DATA_BLOCK "DI_SYSTEM_STRING_NAMES_ENG"
{ S7_Optimized_Access := 'FALSE' }
VERSION : 0.1
NON_RETAIN
"DT_DI_STRING_SYSTEM_NAMES"

BEGIN
   NUM[0] := 'Unit control and prot. +1CJA01';
   NUM[1] := 'Unit control and prot. +1CJA01';
   NUM[2] := 'Unit control and prot. +1CJA01';
   NUM[3] := 'Unit control and prot. +1CJA01';
   NUM[4] := 'Unit control and prot. +1CJA01';
   NUM[5] := 'Unit control and prot. +1CJA01';
   NUM[6] := 'Unit control and prot. +1CJA01';
   NUM[7] := 'Power house pushbutton ';
   NUM[8] := 'Unit control and prot. +1CJA01';
   NUM[9] := '';
   NUM[10] := 'Unit control and prot. +1CJA01';
   NUM[11] := 'Unit control and prot. +1CJA01';
   NUM[12] := 'Unit control and prot. +1CJA01';
   NUM[13] := 'Unit control and prot. +1CJA01';
   NUM[14] := 'Unit control and prot. +1CJA01';
   NUM[15] := '';
   NUM[16] := '';
   NUM[17] := 'Unit GCB cubicle +BAC01';
   NUM[18] := 'Unit GCB cubicle +BAC01';
   NUM[19] := 'Unit GCB cubicle +BAC01';
   NUM[20] := 'Unit GCB cubicle +BAC01';
   NUM[21] := '';
   NUM[22] := '';
   NUM[23] := 'Unit GCB cubicle +BAC01';
   NUM[24] := 'Unit GCB cubicle +BAC01';
   NUM[25] := 'Unit control and prot. +1CJA01';
   NUM[26] := '';
   NUM[27] := '';
   NUM[28] := 'Unit control and prot. +1CJA01';
   NUM[29] := '';
   NUM[30] := 'Unit GCB cubicle +BAC01';
   NUM[31] := 'Common control and prot. +0CJA01';
   NUM[32] := '';
   NUM[33] := '';
   NUM[34] := 'Auxiliary supply cubicle +0BFA01';
   NUM[35] := '';
   NUM[36] := 'Unit Aux. Power Supply +BFA01';
   NUM[37] := '';
   NUM[38] := '';
   NUM[39] := '';
   NUM[40] := '';
   NUM[41] := '';
   NUM[42] := '';
   NUM[43] := '';
   NUM[44] := '';
   NUM[45] := '';
   NUM[46] := '';
   NUM[47] := 'Unit Aux. Power Supply +BFA01';
   NUM[48] := '';
   NUM[49] := 'Unit Aux. Power Supply +BFA01';
   NUM[50] := 'Unit Aux. Power Supply +BFA01';
   NUM[51] := 'Unit Aux. Power Supply +BFA01';
   NUM[52] := '';
   NUM[53] := 'Unit Aux. Power Supply +BFA01';
   NUM[54] := '';
   NUM[55] := '';
   NUM[56] := 'Unit Aux. Power Supply +BFA01';
   NUM[57] := '';
   NUM[58] := 'Unit Aux. Power Supply +BFA01';
   NUM[59] := 'Unit Aux. Power Supply +BFA01';
   NUM[60] := 'Unit Aux. Power Supply +BFA01';
   NUM[61] := 'Unit Aux. Power Supply +BFA01';
   NUM[62] := 'Unit Aux. Power Supply +BFA01';
   NUM[63] := '';
   NUM[64] := '';
   NUM[65] := '';
   NUM[66] := '';
   NUM[67] := '';
   NUM[68] := 'Unit GCB cubicle +BAC01';
   NUM[69] := 'Unit GCB cubicle +BAC01';
   NUM[70] := '';
   NUM[71] := '';
   NUM[72] := '';
   NUM[73] := '';
   NUM[74] := 'Unit GCB cubicle +BAC01';
   NUM[75] := '';
   NUM[76] := '';
   NUM[77] := '';
   NUM[78] := '';
   NUM[79] := '';
   NUM[80] := '';
   NUM[81] := '';
   NUM[82] := '';
   NUM[83] := 'Unit GCB cubicle +BAC01';
   NUM[84] := '';
   NUM[85] := '';
   NUM[86] := 'Unit GCB cubicle +BAC01';
   NUM[87] := '';
   NUM[88] := '';
   NUM[89] := '';
   NUM[90] := '';
   NUM[91] := '';
   NUM[92] := '';
   NUM[93] := '';
   NUM[94] := '';
   NUM[95] := '';
   NUM[96] := '';
   NUM[97] := '';
   NUM[98] := '';
   NUM[99] := 'Unit control and prot. +1CJA01';
   NUM[100] := 'Unit control and prot. +1CJA01';
   NUM[101] := '';
   NUM[102] := '';
   NUM[103] := '';
   NUM[104] := '';
   NUM[105] := '';
   NUM[106] := '';
   NUM[107] := '';
   NUM[108] := '';
   NUM[109] := '';
   NUM[110] := '';
   NUM[111] := '';
   NUM[112] := '';
   NUM[113] := 'Unit Generator - 1MKA10';
   NUM[114] := 'Unit Generator - 1MKA10';
   NUM[115] := '';
   NUM[116] := '';
   NUM[117] := '';
   NUM[118] := '';
   NUM[119] := '';
   NUM[120] := '';
   NUM[121] := '';
   NUM[122] := '';
   NUM[123] := '';
   NUM[124] := '';
   NUM[125] := '';
   NUM[126] := '';
   NUM[127] := '';
   NUM[128] := 'Unit GCB cubicle +BAC01';
   NUM[129] := '';
   NUM[130] := 'Unit GCB cubicle +BAC01';
   NUM[131] := 'Unit GCB cubicle +BAC01';
   NUM[132] := '';
   NUM[133] := '';
   NUM[134] := '';
   NUM[135] := '';
   NUM[136] := '';
   NUM[137] := '';
   NUM[138] := '';
   NUM[139] := '';
   NUM[140] := 'AJA03 - Transformator fedder';
   NUM[141] := '';
   NUM[142] := '';
   NUM[143] := '';
   NUM[144] := '';
   NUM[145] := '';
   NUM[146] := '';
   NUM[147] := '';
   NUM[148] := '';
   NUM[149] := '';
   NUM[150] := '';
   NUM[151] := '';
   NUM[152] := '';
   NUM[153] := '';
   NUM[154] := '';
   NUM[155] := '';
   NUM[156] := '';
   NUM[157] := '';
   NUM[158] := '';
   NUM[159] := '';
   NUM[160] := '';
   NUM[161] := '';
   NUM[162] := '';
   NUM[163] := '';
   NUM[164] := '';
   NUM[165] := '';
   NUM[166] := '';
   NUM[167] := '';
   NUM[168] := '';
   NUM[169] := '';
   NUM[170] := '';
   NUM[171] := '';
   NUM[172] := '';
   NUM[173] := '';
   NUM[174] := '';
   NUM[175] := '';
   NUM[176] := '';
   NUM[177] := '';
   NUM[178] := '';
   NUM[179] := '';
   NUM[180] := '';
   NUM[181] := '';
   NUM[182] := '';
   NUM[183] := '';
   NUM[184] := '';
   NUM[185] := '';
   NUM[186] := '';
   NUM[187] := '';
   NUM[188] := '';
   NUM[189] := '';
   NUM[190] := '';
   NUM[191] := '';
   NUM[192] := 'Unit MIV +1MEA10';
   NUM[193] := '';
   NUM[194] := 'Unit MIV +1MEA10';
   NUM[195] := '';
   NUM[196] := '';
   NUM[197] := '';
   NUM[198] := '';
   NUM[199] := '';
   NUM[200] := '';
   NUM[201] := 'Unit Turbine +1MEA10';
   NUM[202] := 'Unit Turbine +1MEA10';
   NUM[203] := 'Unit control and prot. +1CJA01';
   NUM[204] := '';
   NUM[205] := '';
   NUM[206] := 'Unit control and prot. +1CJA01';
   NUM[207] := 'Unit control and prot. +1CJA01';
   NUM[208] := 'Unit control and prot. +1CJA01';
   NUM[209] := '';
   NUM[210] := '';
   NUM[211] := '';
   NUM[212] := '';
   NUM[213] := '';
   NUM[214] := '';
   NUM[215] := '';
   NUM[216] := '';
   NUM[217] := '';
   NUM[218] := '';
   NUM[219] := '';
   NUM[220] := '';
   NUM[221] := '';
   NUM[222] := '';
   NUM[223] := '';
   NUM[224] := '';
   NUM[225] := 'Unit HPU +1MEX10';
   NUM[226] := '';
   NUM[227] := '';
   NUM[228] := 'Unit HPU +1MEX10';
   NUM[229] := '';
   NUM[230] := '';
   NUM[231] := '';
   NUM[232] := '';
   NUM[233] := 'Unit HPU +1MEX10';
   NUM[234] := 'Unit HPU +1MEX10';
   NUM[235] := '';
   NUM[236] := '';
   NUM[237] := 'Unit HPU +1MEX10';
   NUM[238] := 'Unit HPU +1MEX10';
   NUM[239] := '';
   NUM[240] := '';
   NUM[241] := '';
   NUM[242] := 'Unit control and prot. +1CJA01';
   NUM[243] := 'Unit control and prot. +1CJA01';
   NUM[244] := '';
   NUM[245] := 'HPU +1MEX10';
   NUM[246] := '';
   NUM[247] := '';
   NUM[248] := '';
   NUM[249] := '';
   NUM[250] := '';
   NUM[251] := '';
   NUM[252] := '';
   NUM[253] := '';
   NUM[254] := '';
   NUM[255] := '';
   NUM[256] := '';
   NUM[257] := '';
   NUM[258] := '';
   NUM[259] := 'Unit control and prot. +1CJA01';
   NUM[260] := 'Unit control and prot. +1CJA01';
   NUM[261] := '';
   NUM[262] := '';
   NUM[263] := '';
   NUM[264] := 'Unit control and prot. +1CJA01';
   NUM[265] := 'Unit control and prot. +1CJA01';
   NUM[266] := '';
   NUM[267] := '';
   NUM[268] := '';
   NUM[269] := '';
   NUM[270] := '';
   NUM[271] := '';
   NUM[272] := '';
   NUM[273] := '';
   NUM[274] := '';
   NUM[275] := '';
   NUM[276] := '';
   NUM[277] := '';
   NUM[278] := '';
   NUM[279] := '';
   NUM[280] := '';
   NUM[281] := '';
   NUM[282] := '';
   NUM[283] := '';
   NUM[284] := '';
   NUM[285] := '';
   NUM[286] := '';
   NUM[287] := '';
   NUM[288] := '';
   NUM[289] := '';
   NUM[290] := '';
   NUM[291] := '';
   NUM[292] := '';
   NUM[293] := '';
   NUM[294] := '';
   NUM[295] := '';
   NUM[296] := '';
   NUM[297] := '';
   NUM[298] := '';
   NUM[299] := '';
   NUM[300] := '';
   NUM[301] := '';
   NUM[302] := '';
   NUM[303] := '';
   NUM[304] := '';
   NUM[305] := '';
   NUM[306] := '';
   NUM[307] := '';
   NUM[308] := '';
   NUM[309] := '';
   NUM[310] := '';
   NUM[311] := '';
   NUM[312] := '';
   NUM[313] := '';
   NUM[314] := '';
   NUM[315] := '';
   NUM[316] := '';
   NUM[317] := '';
   NUM[318] := '';
   NUM[319] := '';
   NUM[320] := '';
   NUM[321] := '';
   NUM[322] := '';
   NUM[323] := '';
   NUM[324] := '';
   NUM[325] := '';
   NUM[326] := '';
   NUM[327] := '';
   NUM[328] := '';
   NUM[329] := '';
   NUM[330] := '';
   NUM[331] := '';
   NUM[332] := '';
   NUM[333] := '';
   NUM[334] := '';
   NUM[335] := '';
   NUM[336] := '';
   NUM[337] := '';
   NUM[338] := '';
   NUM[339] := '';
   NUM[340] := '';
   NUM[341] := '';
   NUM[342] := '';
   NUM[343] := '';
   NUM[344] := '';
   NUM[345] := '';
   NUM[346] := '';
   NUM[347] := '';
   NUM[348] := '';
   NUM[349] := '';
   NUM[350] := '';
   NUM[351] := '';
   NUM[352] := 'Unit Turbine +1MEA10';
   NUM[353] := '';
   NUM[354] := '';
   NUM[355] := '';
   NUM[356] := '';
   NUM[357] := '';
   NUM[358] := '';
   NUM[359] := '';
   NUM[360] := '';
   NUM[361] := '';
   NUM[362] := '';
   NUM[363] := '';
   NUM[364] := '';
   NUM[365] := '';
   NUM[366] := '';
   NUM[367] := '';
   NUM[368] := '';
   NUM[369] := '';
   NUM[370] := '';
   NUM[371] := '';
   NUM[372] := '';
   NUM[373] := '';
   NUM[374] := '';
   NUM[375] := '';
   NUM[376] := '';
   NUM[377] := '';
   NUM[378] := '';
   NUM[379] := '';
   NUM[380] := '';
   NUM[381] := '';
   NUM[382] := '';
   NUM[383] := '';
   NUM[384] := 'Unit TRAFO +0BAT01';
   NUM[385] := 'Unit TRAFO +0BAT01';
   NUM[386] := 'Unit TRAFO +0BAT01';
   NUM[387] := 'Unit TRAFO +0BAT01';
   NUM[388] := '';
   NUM[389] := '';
   NUM[390] := '';
   NUM[391] := '';
   NUM[392] := 'Unit SS TRAFO +1BFT01';
   NUM[393] := 'Unit SS TRAFO +1BFT01';
   NUM[394] := 'Unit SS TRAFO +1BFT01';
   NUM[395] := 'Unit SS TRAFO +1BFT01';
   NUM[396] := '';
   NUM[397] := '';
   NUM[398] := '';
   NUM[399] := '';
   NUM[400] := '';
   NUM[401] := '';
   NUM[402] := '';
   NUM[403] := '';
   NUM[404] := '';
   NUM[405] := '';
   NUM[406] := '';
   NUM[407] := '';
   NUM[408] := '';
   NUM[409] := '';
   NUM[410] := '';
   NUM[411] := '';
   NUM[412] := '';
   NUM[413] := '';
   NUM[414] := '';
   NUM[415] := '';
   NUM[416] := '';
   NUM[417] := '';
   NUM[418] := '';
   NUM[419] := '';
   NUM[420] := '';
   NUM[421] := '';
   NUM[422] := '';
   NUM[423] := '';
   NUM[424] := '';
   NUM[425] := '';
   NUM[426] := '';
   NUM[427] := '';
   NUM[428] := '';
   NUM[429] := '';
   NUM[430] := '';
   NUM[431] := '';
   NUM[432] := '';
   NUM[433] := '';
   NUM[434] := '';
   NUM[435] := '';
   NUM[436] := '';
   NUM[437] := '';
   NUM[438] := '';
   NUM[439] := '';
   NUM[440] := '';
   NUM[441] := '';
   NUM[442] := '';
   NUM[443] := '';
   NUM[444] := '';
   NUM[445] := '';
   NUM[446] := '';
   NUM[447] := '';
   NUM[448] := 'Unit control and prot. +1CJA01';
   NUM[449] := 'Unit GCB cubicle +BAC01';
   NUM[450] := 'Unit GCB cubicle +BAC01';
   NUM[451] := 'Unit control and prot. +1CJA01';
   NUM[452] := 'Unit control and prot. +1CJA01';
   NUM[453] := '';
   NUM[454] := '';
   NUM[455] := '';
   NUM[456] := '';
   NUM[457] := 'Unit control and prot. +1CJA01';
   NUM[458] := '';
   NUM[459] := '';
   NUM[460] := 'Unit control and prot. +1CJA01';
   NUM[461] := '';
   NUM[462] := 'Unit control and prot. +1CJA01';
   NUM[463] := 'Unit control and prot. +1CJA01';
   NUM[464] := 'Unit control and prot. +1CJA01';
   NUM[465] := 'Unit control and prot. +1CJA01';
   NUM[466] := 'Unit Generator - 1MKA10';
   NUM[467] := 'Unit Generator - 1MKA10';
   NUM[468] := 'Unit Generator - 1MKA10';
   NUM[469] := '';
   NUM[470] := '';
   NUM[471] := '';
   NUM[472] := '';
   NUM[473] := '';
   NUM[474] := '';
   NUM[475] := '';
   NUM[476] := '';
   NUM[477] := '';
   NUM[478] := '';
   NUM[479] := 'Unit Generator - 1MKA10';
   NUM[480] := 'MV Cubicle - AJA04';
   NUM[481] := 'MV Cubicle - AJA04';
   NUM[482] := '';
   NUM[483] := '';
   NUM[484] := 'MV Cubicle - AJA04';
   NUM[485] := '';
   NUM[486] := '';
   NUM[487] := '';
   NUM[488] := '';
   NUM[489] := '';
   NUM[490] := '';
   NUM[491] := '';
   NUM[492] := '';
   NUM[493] := '';
   NUM[494] := '';
   NUM[495] := '';
   NUM[496] := '';
   NUM[497] := '';
   NUM[498] := '';
   NUM[499] := '';
   NUM[500] := '';
   NUM[501] := '';
   NUM[502] := '';
   NUM[503] := '';
   NUM[504] := '';
   NUM[505] := '';
   NUM[506] := '';
   NUM[507] := '';
   NUM[508] := '';
   NUM[509] := '';
   NUM[510] := '';
   NUM[511] := '';
   NUM[512] := 'MV Cubicle - AJA03';
   NUM[513] := 'MV Cubicle - AJA03';
   NUM[514] := '';
   NUM[515] := 'MV Cubicle - AJA03';
   NUM[516] := 'MV Cubicle - AJA03';
   NUM[517] := '';
   NUM[518] := '';
   NUM[519] := '';
   NUM[520] := '';
   NUM[521] := '';
   NUM[522] := 'MV Cubicle - AJA03';
   NUM[523] := 'MV Cubicle - AJA03';
   NUM[524] := '';
   NUM[525] := '';
   NUM[526] := 'MV Cubicle - AJA03';
   NUM[527] := '';
   NUM[528] := '';
   NUM[529] := '';
   NUM[530] := 'MV Cubicle - AJA04';
   NUM[531] := 'MV Cubicle - AJA03';
   NUM[532] := '';
   NUM[533] := '';
   NUM[534] := '';
   NUM[535] := 'MV Cubicle - AJA03';
   NUM[536] := 'MV Cubicle - AJA03';
   NUM[537] := '';
   NUM[538] := '';
   NUM[539] := '';
   NUM[540] := '';
   NUM[541] := '';
   NUM[542] := 'MV Cubicle - AJA03';
   NUM[543] := 'MV Cubicle - AJA04';
   NUM[544] := '';
   NUM[545] := '';
   NUM[546] := '';
   NUM[547] := '';
   NUM[548] := '';
   NUM[549] := '';
   NUM[550] := '';
   NUM[551] := '';
   NUM[552] := '';
   NUM[553] := '';
   NUM[554] := '';
   NUM[555] := '';
   NUM[556] := '';
   NUM[557] := '';
   NUM[558] := '';
   NUM[559] := '';
   NUM[560] := '';
   NUM[561] := '';
   NUM[562] := '';
   NUM[563] := '';
   NUM[564] := '';
   NUM[565] := '';
   NUM[566] := '';
   NUM[567] := '';
   NUM[568] := '';
   NUM[569] := '';
   NUM[570] := '';
   NUM[571] := '';
   NUM[572] := '';
   NUM[573] := '';
   NUM[574] := '';
   NUM[575] := '';
   NUM[576] := '';
   NUM[577] := '';
   NUM[578] := '';
   NUM[579] := '';
   NUM[580] := '';
   NUM[581] := '';
   NUM[582] := '';
   NUM[583] := '';
   NUM[584] := '';
   NUM[585] := '';
   NUM[586] := '';
   NUM[587] := '';
   NUM[588] := '';
   NUM[589] := '';
   NUM[590] := '';
   NUM[591] := '';
   NUM[592] := '';
   NUM[593] := '';
   NUM[594] := '';
   NUM[595] := '';
   NUM[596] := '';
   NUM[597] := '';
   NUM[598] := '';
   NUM[599] := '';
   NUM[600] := '';
   NUM[601] := '';
   NUM[602] := '';
   NUM[603] := '';
   NUM[604] := '';
   NUM[605] := '';
   NUM[606] := '';
   NUM[607] := 'Unit 1 control and prot. +1CJA01';

END_DATA_BLOCK
DATA_BLOCK "DI_STRING_NAMES_ENG"
{ S7_Optimized_Access := 'FALSE' }
VERSION : 0.1
NON_RETAIN
"DT_DI_STRING_NAMES"

BEGIN
   NUM[0] := 'Maintance switch active (-S100)';
   NUM[1] := 'Local control active (-S103)';
   NUM[2] := 'Auto control active (-S104)';
   NUM[3] := 'Start pushbutton pressed (-S210)';
   NUM[4] := 'Stop pushbutton not pressed (-S211)';
   NUM[5] := 'Reset Alarms (-S302)';
   NUM[6] := 'ESD pushbutton not pressed (-S301)';
   NUM[7] := 'External ESD pushbutton  not pressed';
   NUM[8] := 'ESD relay OK (-K301)';
   NUM[9] := 'Watchdog active';
   NUM[10] := 'External Signals PS OK (-F36, 1K28)';
   NUM[11] := 'DC MCB group alarm (-F41)';
   NUM[12] := 'DC MCB group trip (-F34, -F37, -F38, -F39)';
   NUM[13] := 'Synchronization manual';
   NUM[14] := 'Synchronization auto';
   NUM[15] := 'Synchronization start';
   NUM[16] := 'Synchronization stop';
   NUM[17] := 'Synchronizer MCB OK (-F26)';
   NUM[18] := 'Synchronization active / Contactor closed (-K1)';
   NUM[19] := 'Synchronization speed down (-F25G)';
   NUM[20] := 'Synchronization speed up (-F25G)';
   NUM[21] := 'GCB switch ON pushbutton';
   NUM[22] := 'GCB switch OFF pushbutton';
   NUM[23] := 'GCB closed (-Q1)';
   NUM[24] := 'GCB open (-Q1)';
   NUM[25] := 'Generator overspeed Trip (-K311) ';
   NUM[26] := 'Remote start';
   NUM[27] := 'Remote stop';
   NUM[28] := 'Quick shutdown relay OK (-K401)';
   NUM[29] := 'Remote reset';
   NUM[30] := 'Synchroscope contactor closed (-K1)';
   NUM[31] := 'Trip from Common to Unit 1 (-2K01)';
   NUM[32] := 'AC MCBs group alarm OK';
   NUM[33] := 'AC MCBs group trip OK';
   NUM[34] := 'DC MCB group alarm (-F31,-F422)';
   NUM[35] := 'DC MCB group trip (-F38,39,40,44,45)';
   NUM[36] := 'Main CB ON (-Q0)';
   NUM[37] := 'Main CB OFF';
   NUM[38] := 'Main CB manual';
   NUM[39] := 'Main CB autopmatic';
   NUM[40] := 'Main CB tripped';
   NUM[41] := 'Diesel CB ON';
   NUM[42] := 'Diesel CB OFF';
   NUM[43] := 'Diesel CB manual';
   NUM[44] := 'Diesel CB automatic';
   NUM[45] := 'Overspeed protection MCB OK';
   NUM[46] := 'AC voltage OK (-F411, -K411)';
   NUM[47] := 'Voltage before Main CB OK (-F411, -K411)';
   NUM[48] := 'Voltage before Diesel CB OK';
   NUM[49] := 'Surge arrestor OK (-FU1)';
   NUM[50] := 'AC/DC rectifier 1 OK (-F80, -U101)';
   NUM[51] := 'AC/DC rectifier 2 OK (-F81, -U102)';
   NUM[52] := 'AC/DC rectifier 3 OK';
   NUM[53] := 'Battery connected (-FB, -F421, -K201)';
   NUM[54] := 'Common DC power supply OK (-F0)';
   NUM[55] := 'Intake cubicle AC suppy MCB ON (-F7)';
   NUM[56] := 'Unit (+1CJA01) Cubicle AC Power Supply OK (-F71)';
   NUM[57] := 'Powerhouse distribution panel MCB closed (-F5)';
   NUM[58] := 'Workstation UPS MCB OK (-F32)';
   NUM[59] := 'Unit (+1CJA01) Cubicle DC Power Supply OK (-F10)';
   NUM[60] := 'GCB (+BAC01) Cubicle DC Power Suppy OK (-F11)';
   NUM[61] := 'MV Cubicle DC Power Suppy OK (-F12)';
   NUM[62] := 'MV Cubicle AC Power Suppy OK  (-F83)';
   NUM[63] := 'Common DC power supply (-F0)';
   NUM[64] := 'Spare 64';
   NUM[65] := 'Spare 65';
   NUM[66] := 'Spare 66';
   NUM[67] := 'Spare 67';
   NUM[68] := 'Grid VT Meas MCB OK (-F51, -F52)';
   NUM[69] := 'Gen. VT Meas. MCB OK (-F53)';
   NUM[70] := 'Spare 70';
   NUM[71] := 'Spare 71';
   NUM[72] := 'Spare 72';
   NUM[73] := 'Spare 73';
   NUM[74] := 'GCB ready for close (-Q1)';
   NUM[75] := 'Spare 75';
   NUM[76] := 'GCB spring charged (-Q1)';
   NUM[77] := 'Spare 77';
   NUM[78] := 'Generator CB control MCB ON (-F62)';
   NUM[79] := 'Spare 79';
   NUM[80] := 'Spare 80';
   NUM[81] := 'Spare 81';
   NUM[82] := 'Spare 82';
   NUM[83] := 'Surge Arrester OK (-F60, -FU1)';
   NUM[84] := 'Spare 84';
   NUM[85] := 'Spare 85';
   NUM[86] := 'DC MCB Group Trip (-F4, -F7, -F11, -F14)';
   NUM[87] := 'Aux transformer supply switch ON (-Q2)';
   NUM[88] := 'Spare 88';
   NUM[89] := 'Surge arrestor 2 OK (-F61, -FU2)';
   NUM[90] := 'Spare 90';
   NUM[91] := 'Spare 91';
   NUM[92] := 'Spare 92';
   NUM[93] := 'Spare 93';
   NUM[94] := 'Spare 94';
   NUM[95] := 'Lamp Test (-S203)';
   NUM[96] := 'Generator voltage meas';
   NUM[97] := 'Spare';
   NUM[98] := 'Spare';
   NUM[99] := 'Generator heater CB ON (-F56)';
   NUM[100] := 'Generator heater contactor closed (-K56)';
   NUM[101] := 'Spare';
   NUM[102] := 'Spare';
   NUM[103] := 'Spare';
   NUM[104] := 'Spare';
   NUM[105] := 'Spare';
   NUM[106] := 'Spare';
   NUM[107] := 'Spare';
   NUM[108] := 'Spare';
   NUM[109] := 'Spare';
   NUM[110] := 'Generator lubrication oil level min';
   NUM[111] := 'Generator greasing pump ON (-SG24)';
   NUM[112] := 'Generator Vibration Trip (-VSE002)';
   NUM[113] := '+1MKA10 Generator Oil Level High (1CJA01 -1K05)';
   NUM[114] := '+1MKA10 Generator Oil Level Too High (1CJA01 -1K';
   NUM[115] := 'Spare';
   NUM[116] := 'Spare';
   NUM[117] := 'Spare';
   NUM[118] := 'Spare';
   NUM[119] := 'Spare';
   NUM[120] := 'Spare';
   NUM[121] := 'Spare';
   NUM[122] := 'Spare';
   NUM[123] := 'Spare';
   NUM[124] := 'Spare';
   NUM[125] := 'Spare';
   NUM[126] := 'Spare';
   NUM[127] := 'Spare';
   NUM[128] := 'Generator Protection Trip (-F311)';
   NUM[129] := 'Spare';
   NUM[130] := 'Generator Protection Alarm (-F311)';
   NUM[131] := 'Generator Protection Live (-F311)';
   NUM[132] := 'Spare';
   NUM[133] := 'Spare';
   NUM[134] := 'Spare';
   NUM[135] := 'Spare';
   NUM[136] := 'Spare';
   NUM[137] := 'Spare';
   NUM[138] := 'Spare';
   NUM[139] := 'Spare';
   NUM[140] := 'AJA03 -Line protection trip 1 (-REF615)';
   NUM[141] := 'AJA04 -Line protection trip 2 (-F200)';
   NUM[142] := 'AJA04 - Line protection alarm (-F200)';
   NUM[143] := 'AKA04 - Line protection live (-F200)';
   NUM[144] := 'Spare';
   NUM[145] := 'Spare';
   NUM[146] := 'Spare';
   NUM[147] := 'Spare';
   NUM[148] := 'Spare';
   NUM[149] := 'Spare';
   NUM[150] := 'Spare';
   NUM[151] := 'Spare';
   NUM[152] := 'Spare';
   NUM[153] := 'Spare';
   NUM[154] := 'Spare';
   NUM[155] := 'Spare';
   NUM[156] := 'Spare';
   NUM[157] := 'Spare';
   NUM[158] := 'Spare';
   NUM[159] := 'Spare';
   NUM[160] := 'Surge arrestor OK (-FU1)';
   NUM[161] := 'Incoming supply CB ON (-Q1)';
   NUM[162] := 'Rectifier OK (-F3)';
   NUM[163] := 'DC MCB ok group alarm (-F31, -F40)';
   NUM[164] := 'AC MCB ok group alarm (-F2,-F5,-F6)';
   NUM[165] := 'PSU (-U101) - ALARM';
   NUM[166] := 'PSU (-U101) - Battery mode';
   NUM[167] := 'PSU (-U101) - Charge mode';
   NUM[168] := 'Spare';
   NUM[169] := 'Spare';
   NUM[170] := 'Spare';
   NUM[171] := 'Spare';
   NUM[172] := 'Spare';
   NUM[173] := 'Spare';
   NUM[174] := 'Spare';
   NUM[175] := 'Spare';
   NUM[176] := 'Spare';
   NUM[177] := 'Spare';
   NUM[178] := 'Spare';
   NUM[179] := 'Spare';
   NUM[180] := 'Spare';
   NUM[181] := 'Spare';
   NUM[182] := 'Spare';
   NUM[183] := 'Spare';
   NUM[184] := 'Spare';
   NUM[185] := 'Spare';
   NUM[186] := 'Spare';
   NUM[187] := 'Spare';
   NUM[188] := 'Spare';
   NUM[189] := 'Spare';
   NUM[190] := 'Spare';
   NUM[191] := 'Spare';
   NUM[192] := 'MIV closed (+1CJA01 -1K33)';
   NUM[193] := 'Spare';
   NUM[194] := 'MIV open (+1CJA01 -1K32)';
   NUM[195] := 'Spare';
   NUM[196] := 'Spare';
   NUM[197] := 'MIV CB closed (-F52)';
   NUM[198] := 'MIV contactor closed (-K52, -K53)';
   NUM[199] := 'MIV heater MCB closed (-F58)';
   NUM[200] := 'Spare';
   NUM[201] := 'Bypass OPEN (ARCON, +1CJA10 -1K07)';
   NUM[202] := 'Bypass CLOSED (-ARCON, +1CJA10 -1K08)';
   NUM[203] := 'Bypass MCB ON (-F40)';
   NUM[204] := 'Spare';
   NUM[205] := 'Bypass contactor closed (-K101)';
   NUM[206] := 'Bypass opening contactor closed (-K102)';
   NUM[207] := 'Bypass closing contactor ON (-K101)';
   NUM[208] := 'Bypass torque swtich (O/C) (-K206)';
   NUM[209] := 'Spare';
   NUM[210] := 'Spare';
   NUM[211] := 'Spare';
   NUM[212] := 'Spare';
   NUM[213] := 'Spare';
   NUM[214] := 'MIV Torque-switch closed (-1K06)';
   NUM[215] := 'MIV Torque-switch open (-1K05)';
   NUM[216] := 'MIV Thermoswitch (-1K13)';
   NUM[217] := 'Spare';
   NUM[218] := 'Spare';
   NUM[219] := 'Spare';
   NUM[220] := 'Spare';
   NUM[221] := 'Spare';
   NUM[222] := 'Spare';
   NUM[223] := 'Spare';
   NUM[224] := 'Spare';
   NUM[225] := 'HPU Filter Clogging Indicator OK (-600S1, +1CJA01 -1K15)';
   NUM[226] := 'Spare';
   NUM[227] := 'Spare';
   NUM[228] := 'Accumulator ESD Pressure OK (-IFM, +1CJA01 -1K31)';
   NUM[229] := 'HPU min';
   NUM[230] := 'HPU max';
   NUM[231] := 'Accumulator start/stop pump (-X3';
   NUM[232] := 'System pressure OK (-640B4)';
   NUM[233] := 'HPU Oil Level Too Low (1MEX10 -640B2, 1CJA01 -1K';
   NUM[234] := 'HPU Oil Level Low (1MEX10 -640B2, 1CJA01 -1K12) ';
   NUM[235] := 'Spare';
   NUM[236] := '';
   NUM[237] := 'HPU Oil Temperature High (-640B1, +1CJA01 - 1K13';
   NUM[238] := 'HPU Oil Temperature Too High (-640B1, +1CJA01 - ';
   NUM[239] := 'Spare';
   NUM[240] := 'Spare';
   NUM[241] := 'Spare';
   NUM[242] := 'HPU heater CB ON (-F57)';
   NUM[243] := 'HPU heater contactor closed (-K57)';
   NUM[244] := 'HPU control MCB closed (-F59)';
   NUM[245] := 'HPU ESD Pushbutton pressed';
   NUM[246] := 'Spare';
   NUM[247] := 'Spare';
   NUM[248] := 'Spare';
   NUM[249] := 'Spare';
   NUM[250] := 'Spare';
   NUM[251] := 'Spare';
   NUM[252] := 'Spare';
   NUM[253] := 'Spare';
   NUM[254] := 'Spare';
   NUM[255] := 'Spare';
   NUM[256] := 'Spare';
   NUM[257] := 'Spare';
   NUM[258] := 'Spare';
   NUM[259] := 'HPU Pump 1 CB ON (-F51)';
   NUM[260] := 'HPU Pump 1 contactor closed (-K51)';
   NUM[261] := 'Spare';
   NUM[262] := 'Spare';
   NUM[263] := 'Spare';
   NUM[264] := 'HPU Pump 2 CB ON (-F52)';
   NUM[265] := 'HPU Pump 2 contactor closed (-K52)';
   NUM[266] := 'Spare';
   NUM[267] := 'Spare';
   NUM[268] := 'Spare';
   NUM[269] := 'Spare';
   NUM[270] := 'Spare';
   NUM[271] := 'Spare';
   NUM[272] := 'Spare';
   NUM[273] := 'Spare';
   NUM[274] := 'Spare';
   NUM[275] := 'Spare';
   NUM[276] := 'Spare';
   NUM[277] := 'Spare';
   NUM[278] := 'Spare';
   NUM[279] := 'Spare';
   NUM[280] := 'Spare';
   NUM[281] := 'Spare';
   NUM[282] := 'Spare';
   NUM[283] := 'Spare';
   NUM[284] := 'Spare';
   NUM[285] := 'Spare';
   NUM[286] := 'Spare';
   NUM[287] := 'Spare';
   NUM[288] := 'Spare';
   NUM[289] := 'Spare';
   NUM[290] := 'Spare';
   NUM[291] := 'Spare';
   NUM[292] := 'Spare';
   NUM[293] := 'Spare';
   NUM[294] := 'Spare';
   NUM[295] := 'Spare';
   NUM[296] := 'Spare';
   NUM[297] := 'Spare';
   NUM[298] := 'Spare';
   NUM[299] := 'Spare';
   NUM[300] := 'Spare';
   NUM[301] := 'Spare';
   NUM[302] := 'Spare';
   NUM[303] := 'Spare';
   NUM[304] := 'Spare';
   NUM[305] := 'Spare';
   NUM[306] := 'Spare';
   NUM[307] := 'Spare';
   NUM[308] := 'Spare';
   NUM[309] := 'Spare';
   NUM[310] := 'Spare';
   NUM[311] := 'Spare';
   NUM[312] := 'Spare';
   NUM[313] := 'Spare';
   NUM[314] := 'Spare';
   NUM[315] := 'Spare';
   NUM[316] := 'Spare';
   NUM[317] := 'Spare';
   NUM[318] := 'Spare';
   NUM[319] := 'Spare';
   NUM[320] := 'Spare';
   NUM[321] := 'Spare';
   NUM[322] := 'Spare';
   NUM[323] := 'Spare';
   NUM[324] := 'Spare';
   NUM[325] := 'Spare';
   NUM[326] := 'Spare';
   NUM[327] := 'Spare';
   NUM[328] := 'Spare';
   NUM[329] := 'Spare';
   NUM[330] := 'Spare';
   NUM[331] := 'Spare';
   NUM[332] := 'Spare';
   NUM[333] := 'Spare';
   NUM[334] := 'Spare';
   NUM[335] := 'Spare';
   NUM[336] := 'Spare';
   NUM[337] := 'Spare';
   NUM[338] := 'Spare';
   NUM[339] := 'Spare';
   NUM[340] := 'Spare';
   NUM[341] := 'Spare';
   NUM[342] := 'Spare';
   NUM[343] := 'Spare';
   NUM[344] := 'Spare';
   NUM[345] := 'Spare';
   NUM[346] := 'Spare';
   NUM[347] := 'Spare';
   NUM[348] := 'Spare';
   NUM[349] := 'Spare';
   NUM[350] := 'Spare';
   NUM[351] := 'Spare';
   NUM[352] := 'Wicket gate distortion capture';
   NUM[353] := 'Spare';
   NUM[354] := 'Runner vanes heater MCB ON (-F54)';
   NUM[355] := 'Runner vanes drive cont';
   NUM[356] := 'Runner vanes drive cont';
   NUM[357] := 'Wicket gate heater MCB ON (-F49)';
   NUM[358] := 'Runner vanes drive CB ON (-F51)';
   NUM[359] := 'Wicket gate drive CB ON (-F47)';
   NUM[360] := 'Wicket gate drive cont';
   NUM[361] := 'Wicket gate drive cont';
   NUM[362] := 'Wicket gate heater cont';
   NUM[363] := 'Overspeed trip (turbine) (-K312)';
   NUM[364] := 'Wicket gate torque-switch "C"';
   NUM[365] := 'Wicket gate torque-switch "O"';
   NUM[366] := 'Wicket gate limit-switch "C"';
   NUM[367] := 'Wicket gate limit-switch "O"';
   NUM[368] := 'Runner vanes torque switch "C"';
   NUM[369] := 'Runner vanes torque switch "O"';
   NUM[370] := 'Runner vanes limit switch "C"';
   NUM[371] := 'Runner vanes limit switch "O"';
   NUM[372] := 'Runner vanes thermoswitch (-1K11)';
   NUM[373] := 'Spare';
   NUM[374] := 'Spare';
   NUM[375] := 'Spare';
   NUM[376] := 'Spare';
   NUM[377] := 'Spare';
   NUM[378] := 'Spare';
   NUM[379] := 'Spare';
   NUM[380] := 'Spare';
   NUM[381] := 'Spare';
   NUM[382] := 'Spare';
   NUM[383] := 'Spare';
   NUM[384] := 'Unit trafo - Temperature alarm (+1CJA01 -1K04)';
   NUM[385] := 'Unit trafo - Temperature trip (+1CJA01 -1K03)';
   NUM[386] := 'Unit trafo - Oil level trip (+1CJA01 -1K01)';
   NUM[387] := 'Unit trafo - Pressure trip (+1CJA01 -1K02)';
   NUM[388] := 'Spare';
   NUM[389] := 'Spare';
   NUM[390] := 'Unit trafo - Buchholz alarm';
   NUM[391] := 'Unit trafo 1BAT10 - Gas trip (-1K35)';
   NUM[392] := 'SS Trafo - Oil level Trip (+1CJA01 -1K21)';
   NUM[393] := 'SS Trafo - Pressure Trip (+1CJA01 -1K22)';
   NUM[394] := 'SS Trafo - Temperature Trip (+1CJA01 -1K23)';
   NUM[395] := 'SS Trafo - Temperature Alarm (+1CJA01 -1K24)';
   NUM[396] := 'Spare';
   NUM[397] := 'Spare';
   NUM[398] := 'Spare';
   NUM[399] := 'Spare';
   NUM[400] := 'Spare';
   NUM[401] := 'Spare';
   NUM[402] := 'Spare';
   NUM[403] := 'Spare';
   NUM[404] := 'Spare';
   NUM[405] := 'Spare';
   NUM[406] := 'Spare';
   NUM[407] := 'Spare';
   NUM[408] := 'Spare';
   NUM[409] := 'Spare';
   NUM[410] := 'Spare';
   NUM[411] := 'Spare';
   NUM[412] := 'Spare';
   NUM[413] := 'SS trafo - winding temp U Ok (-TH145)';
   NUM[414] := 'SS trafo - winding temp V Ok (-TH145)';
   NUM[415] := 'SS trafo - winding temp W Ok (-TH145)';
   NUM[416] := 'Spare';
   NUM[417] := 'Spare';
   NUM[418] := 'Spare';
   NUM[419] := 'Spare';
   NUM[420] := 'Spare';
   NUM[421] := 'Spare';
   NUM[422] := 'Spare';
   NUM[423] := 'Spare';
   NUM[424] := 'Spare';
   NUM[425] := 'Spare';
   NUM[426] := 'Spare';
   NUM[427] := 'Spare';
   NUM[428] := 'Spare';
   NUM[429] := 'Spare';
   NUM[430] := 'Spare';
   NUM[431] := 'Spare';
   NUM[432] := 'Spare';
   NUM[433] := 'Spare';
   NUM[434] := 'Spare';
   NUM[435] := 'Spare';
   NUM[436] := 'Spare';
   NUM[437] := 'Spare';
   NUM[438] := 'Spare';
   NUM[439] := 'Spare';
   NUM[440] := 'Spare';
   NUM[441] := 'Spare';
   NUM[442] := 'Spare';
   NUM[443] := 'Spare';
   NUM[444] := 'Spare';
   NUM[445] := 'Spare';
   NUM[446] := 'Spare';
   NUM[447] := 'Spare';
   NUM[448] := 'Excitation contactor closed (-K1)';
   NUM[449] := 'Synchronization Voltage Lower (-F25G)';
   NUM[450] := 'Synchronization Voltage Higher (-F25G)';
   NUM[451] := 'AVR trip (D700-3F -DO7, +1CJA01 -1K37)';
   NUM[452] := 'Excitation device alarm (-DECS 250)';
   NUM[453] := 'Excitation diode monitoring trip (DV0 - RLY3)';
   NUM[454] := 'AVR relay 1';
   NUM[455] := 'AVR relay 2';
   NUM[456] := 'Spare';
   NUM[457] := 'Excitation watchdog OK (-K204)';
   NUM[458] := 'AVR not tripped (-K112)';
   NUM[459] := 'Start AVR ';
   NUM[460] := 'AVR limiter (D700-3F -DO8, +1CJA01 -1K36)';
   NUM[461] := 'Excitation SPARE';
   NUM[462] := 'Excitation AVR active (-DECS 250)';
   NUM[463] := 'Excitation PF ctrl active (-DECS 250)';
   NUM[464] := 'Excitation VAR ctrl active (-DECS 250)';
   NUM[465] := 'Excitation FCR active (-DECS 250)';
   NUM[466] := 'Spare';
   NUM[467] := 'Spare';
   NUM[468] := 'AVR start (D700-3F -DO9, +1CJA01 -1K38)';
   NUM[469] := 'Spare';
   NUM[470] := 'Spare';
   NUM[471] := 'Spare';
   NUM[472] := 'Spare';
   NUM[473] := 'Spare';
   NUM[474] := 'Spare';
   NUM[475] := 'Spare';
   NUM[476] := 'Spare';
   NUM[477] := 'Spare';
   NUM[478] := 'Spare';
   NUM[479] := 'Q1 AREP PS ON (+1CJA01 -1K35)';
   NUM[480] := '0AJA04 - Disconnector closed (-Q2)';
   NUM[481] := '0AJA04 - Disconnector open (-Q2)';
   NUM[482] := 'Spare';
   NUM[483] := '0AJA04 - Earthing switch closed (-Q3)';
   NUM[484] := '0AJA04 - Earthing switch open (-Q3)';
   NUM[485] := '0AKA01 - Voltage detection relay closed (-F23)';
   NUM[486] := '0AKA02 - Voltage trafo MCB closed (-Q11)';
   NUM[487] := '0AKA01 - CB spring charged (-Q0)';
   NUM[488] := 'Spare';
   NUM[489] := '0AKA01 - Remote control (-S60)';
   NUM[490] := '0AKA01 - Cicruit breaker closed (-Q1)';
   NUM[491] := '0AKA01 - Cicruit breaker open (-Q1)';
   NUM[492] := 'Spare';
   NUM[493] := 'Spare';
   NUM[494] := '0AKA01 - DC MCB OK group 1 Trip (-F14)';
   NUM[495] := '0AKA01 - Gas pressure OK (-Q1)';
   NUM[496] := 'Lever inserted';
   NUM[497] := '0AKA01 - 2nd Shunt relase MCB ON (-F5)';
   NUM[498] := 'Spare';
   NUM[499] := '0AKA01 - DC control and signal';
   NUM[500] := '0AKA01 - AC control and signal';
   NUM[501] := '0AKA01 - Charging motor MCB closed (-Q5)';
   NUM[502] := '0AGA02 - Outgoing feeder CB service';
   NUM[503] := '0AKA01 - MV Heaters on (-Q6)';
   NUM[504] := 'Spare';
   NUM[505] := 'Spare';
   NUM[506] := 'Spare';
   NUM[507] := 'Spare';
   NUM[508] := 'Spare';
   NUM[509] := 'Spare';
   NUM[510] := 'Spare';
   NUM[511] := 'Spare';
   NUM[512] := '0AJA03 - Disconnector closed (-S1)';
   NUM[513] := '0AJA03 - Disconnector open (-S1)';
   NUM[514] := 'Spare';
   NUM[515] := '0AJA03 - Earthing switch closed (-PE1)';
   NUM[516] := '0AJA03 - Earthing switch open (-PE1)';
   NUM[517] := '0AKA03 - Voltage present (-F23 -> R1,R2)';
   NUM[518] := 'Spare';
   NUM[519] := 'Spare';
   NUM[520] := 'Spare';
   NUM[521] := 'AJA04 - Local control (-S60)';
   NUM[522] := 'CB Closed (-QL1, -2K10)';
   NUM[523] := 'CB Open (-QL1)';
   NUM[524] := 'Spare';
   NUM[525] := 'Spare';
   NUM[526] := 'DC MCB Group Trip (-F34, -F38)';
   NUM[527] := 'Spare';
   NUM[528] := 'Spare';
   NUM[529] := 'Spare';
   NUM[530] := 'Fuse OK (-BGF1)';
   NUM[531] := 'FUSE Open';
   NUM[532] := 'Spare';
   NUM[533] := 'Spare';
   NUM[534] := 'Spare';
   NUM[535] := 'Breaker FAILURE Trip (-K51)';
   NUM[536] := 'IRF Signal OK (-K201)';
   NUM[537] := 'Control and signal';
   NUM[538] := 'Charging motor MCB closed (-Q5)';
   NUM[539] := 'Spare';
   NUM[540] := '0AKA03 - Voltage trafo MCB closed (-Q11)';
   NUM[541] := 'Spare';
   NUM[542] := 'CB Closed Auxiliary Signal (-QL1) ';
   NUM[543] := 'Fuse Position Open (-BGF1)';
   NUM[544] := 'S';
   NUM[545] := 'S';
   NUM[546] := 'S';
   NUM[547] := 'S';
   NUM[548] := 'S';
   NUM[549] := 'S';
   NUM[550] := 'Spare';
   NUM[551] := 'Spare';
   NUM[552] := 'Spare';
   NUM[553] := 'Spare';
   NUM[554] := 'Spare';
   NUM[555] := 'Spare';
   NUM[556] := 'Spare';
   NUM[557] := 'Spare';
   NUM[558] := 'Spare';
   NUM[559] := 'Spare';
   NUM[560] := 'Spare';
   NUM[561] := 'Spare';
   NUM[562] := 'Spare';
   NUM[563] := 'Spare';
   NUM[564] := 'Spare';
   NUM[565] := 'Spare';
   NUM[566] := 'Spare';
   NUM[567] := 'Spare';
   NUM[568] := 'Spare';
   NUM[569] := 'Spare';
   NUM[570] := 'Spare';
   NUM[571] := 'Spare';
   NUM[572] := 'Spare';
   NUM[573] := 'Spare';
   NUM[574] := 'Spare';
   NUM[575] := 'Spare';
   NUM[576] := '0AKA03 - CB open (-Q1)';
   NUM[577] := '0AKA03 - CB closed (-Q1)';
   NUM[578] := 'Step-up transformer outgoing spring charged';
   NUM[579] := '0AKA03 - ES closed (-Q3)';
   NUM[580] := '0AKA03 - DS open (-Q2)';
   NUM[581] := '0AKA03 - DS closed (-Q2)';
   NUM[582] := 'Step-up transformer outgoing control MCB closed';
   NUM[583] := 'Step-up transf';
   NUM[584] := '0AKA03 - CB closing (-S60)';
   NUM[585] := '0AKA03 - control and signal';
   NUM[586] := '0AKA03 - Charging motor MCB closed (-Q5)';
   NUM[587] := 'Step-up transformer incoming AC MCB closed';
   NUM[588] := '0AKA03 - Voltage trafo MCB closed (-Q11)';
   NUM[589] := '0AGA01 - VT2 MCB closed';
   NUM[590] := '0AGA01 - VT3 MCB closed';
   NUM[591] := '0AKA03 - ES open (-Q3)';
   NUM[592] := '0AKA03 - Voltage detection relay closed (-F23)';
   NUM[593] := 'SPARE';
   NUM[594] := 'SPARE';
   NUM[595] := 'SPARE';
   NUM[596] := 'SPARE';
   NUM[597] := 'SPARE';
   NUM[598] := 'SPARE';
   NUM[599] := 'SPARE';
   NUM[600] := 'SPARE';
   NUM[601] := 'SPARE';
   NUM[602] := 'SPARE';
   NUM[603] := 'SPARE';
   NUM[604] := 'SPARE';
   NUM[605] := 'SPARE';
   NUM[606] := 'SPARE';
   NUM[607] := 'SPARE';

END_DATA_BLOCK
DATA_BLOCK "DI_SYSTEM_STRING_NAMES_GER"
{ S7_Optimized_Access := 'FALSE' }
VERSION : 0.1
NON_RETAIN
"DT_DI_STRING_SYSTEM_NAMES"

BEGIN
   NUM[0] := '';
   NUM[1] := '';
   NUM[2] := '';
   NUM[3] := '';
   NUM[4] := '';
   NUM[5] := '';
   NUM[6] := '';
   NUM[7] := '';
   NUM[8] := '';
   NUM[9] := '';
   NUM[10] := '';
   NUM[11] := '';
   NUM[12] := '';
   NUM[13] := '';
   NUM[14] := '';
   NUM[15] := '';
   NUM[16] := '';
   NUM[17] := '';
   NUM[18] := '';
   NUM[19] := '';
   NUM[20] := '';
   NUM[21] := '';
   NUM[22] := '';
   NUM[23] := '';
   NUM[24] := '';
   NUM[25] := '';
   NUM[26] := '';
   NUM[27] := '';
   NUM[28] := '';
   NUM[29] := '';
   NUM[30] := '';
   NUM[31] := '';
   NUM[32] := '';
   NUM[33] := '';
   NUM[34] := '';
   NUM[35] := '';
   NUM[36] := '';
   NUM[37] := '';
   NUM[38] := '';
   NUM[39] := '';
   NUM[40] := '';
   NUM[41] := '';
   NUM[42] := '';
   NUM[43] := '';
   NUM[44] := '';
   NUM[45] := '';
   NUM[46] := '';
   NUM[47] := '';
   NUM[48] := '';
   NUM[49] := '';
   NUM[50] := '';
   NUM[51] := '';
   NUM[52] := '';
   NUM[53] := '';
   NUM[54] := '';
   NUM[55] := '';
   NUM[56] := '';
   NUM[57] := '';
   NUM[58] := '';
   NUM[59] := '';
   NUM[60] := '';
   NUM[61] := '';
   NUM[62] := '';
   NUM[63] := '';
   NUM[64] := '';
   NUM[65] := '';
   NUM[66] := '';
   NUM[67] := '';
   NUM[68] := '';
   NUM[69] := '';
   NUM[70] := '';
   NUM[71] := '';
   NUM[72] := '';
   NUM[73] := '';
   NUM[74] := '';
   NUM[75] := '';
   NUM[76] := '';
   NUM[77] := '';
   NUM[78] := '';
   NUM[79] := '';
   NUM[80] := '';
   NUM[81] := '';
   NUM[82] := '';
   NUM[83] := '';
   NUM[84] := '';
   NUM[85] := '';
   NUM[86] := '';
   NUM[87] := '';
   NUM[88] := '';
   NUM[89] := '';
   NUM[90] := '';
   NUM[91] := '';
   NUM[92] := '';
   NUM[93] := '';
   NUM[94] := '';
   NUM[95] := '';
   NUM[96] := '';
   NUM[97] := '';
   NUM[98] := '';
   NUM[99] := '';
   NUM[100] := '';
   NUM[101] := '';
   NUM[102] := '';
   NUM[103] := '';
   NUM[104] := '';
   NUM[105] := '';
   NUM[106] := '';
   NUM[107] := '';
   NUM[108] := '';
   NUM[109] := '';
   NUM[110] := '';
   NUM[111] := '';
   NUM[112] := '';
   NUM[113] := '';
   NUM[114] := '';
   NUM[115] := '';
   NUM[116] := '';
   NUM[117] := '';
   NUM[118] := '';
   NUM[119] := '';
   NUM[120] := '';
   NUM[121] := '';
   NUM[122] := '';
   NUM[123] := '';
   NUM[124] := '';
   NUM[125] := '';
   NUM[126] := '';
   NUM[127] := '';
   NUM[128] := '';
   NUM[129] := '';
   NUM[130] := '';
   NUM[131] := '';
   NUM[132] := '';
   NUM[133] := '';
   NUM[134] := '';
   NUM[135] := '';
   NUM[136] := '';
   NUM[137] := '';
   NUM[138] := '';
   NUM[139] := '';
   NUM[140] := '';
   NUM[141] := '';
   NUM[142] := '';
   NUM[143] := '';
   NUM[144] := '';
   NUM[145] := '';
   NUM[146] := '';
   NUM[147] := '';
   NUM[148] := '';
   NUM[149] := '';
   NUM[150] := '';
   NUM[151] := '';
   NUM[152] := '';
   NUM[153] := '';
   NUM[154] := '';
   NUM[155] := '';
   NUM[156] := '';
   NUM[157] := '';
   NUM[158] := '';
   NUM[159] := '';
   NUM[160] := '';
   NUM[161] := '';
   NUM[162] := '';
   NUM[163] := '';
   NUM[164] := '';
   NUM[165] := '';
   NUM[166] := '';
   NUM[167] := '';
   NUM[168] := '';
   NUM[169] := '';
   NUM[170] := '';
   NUM[171] := '';
   NUM[172] := '';
   NUM[173] := '';
   NUM[174] := '';
   NUM[175] := '';
   NUM[176] := '';
   NUM[177] := '';
   NUM[178] := '';
   NUM[179] := '';
   NUM[180] := '';
   NUM[181] := '';
   NUM[182] := '';
   NUM[183] := '';
   NUM[184] := '';
   NUM[185] := '';
   NUM[186] := '';
   NUM[187] := '';
   NUM[188] := '';
   NUM[189] := '';
   NUM[190] := '';
   NUM[191] := '';
   NUM[192] := '';
   NUM[193] := '';
   NUM[194] := '';
   NUM[195] := '';
   NUM[196] := '';
   NUM[197] := '';
   NUM[198] := '';
   NUM[199] := '';
   NUM[200] := '';
   NUM[201] := '';
   NUM[202] := '';
   NUM[203] := '';
   NUM[204] := '';
   NUM[205] := '';
   NUM[206] := '';
   NUM[207] := '';
   NUM[208] := '';
   NUM[209] := '';
   NUM[210] := '';
   NUM[211] := '';
   NUM[212] := '';
   NUM[213] := '';
   NUM[214] := '';
   NUM[215] := '';
   NUM[216] := '';
   NUM[217] := '';
   NUM[218] := '';
   NUM[219] := '';
   NUM[220] := '';
   NUM[221] := '';
   NUM[222] := '';
   NUM[223] := '';
   NUM[224] := '';
   NUM[225] := '';
   NUM[226] := '';
   NUM[227] := '';
   NUM[228] := '';
   NUM[229] := '';
   NUM[230] := '';
   NUM[231] := '';
   NUM[232] := '';
   NUM[233] := '';
   NUM[234] := '';
   NUM[235] := '';
   NUM[236] := '';
   NUM[237] := '';
   NUM[238] := '';
   NUM[239] := '';
   NUM[240] := '';
   NUM[241] := '';
   NUM[242] := '';
   NUM[243] := '';
   NUM[244] := '';
   NUM[245] := '';
   NUM[246] := '';
   NUM[247] := '';
   NUM[248] := '';
   NUM[249] := '';
   NUM[250] := '';
   NUM[251] := '';
   NUM[252] := '';
   NUM[253] := '';
   NUM[254] := '';
   NUM[255] := '';
   NUM[256] := '';
   NUM[257] := '';
   NUM[258] := '';
   NUM[259] := '';
   NUM[260] := '';
   NUM[261] := '';
   NUM[262] := '';
   NUM[263] := '';
   NUM[264] := '';
   NUM[265] := '';
   NUM[266] := '';
   NUM[267] := '';
   NUM[268] := '';
   NUM[269] := '';
   NUM[270] := '';
   NUM[271] := '';
   NUM[272] := '';
   NUM[273] := '';
   NUM[274] := '';
   NUM[275] := '';
   NUM[276] := '';
   NUM[277] := '';
   NUM[278] := '';
   NUM[279] := '';
   NUM[280] := '';
   NUM[281] := '';
   NUM[282] := '';
   NUM[283] := '';
   NUM[284] := '';
   NUM[285] := '';
   NUM[286] := '';
   NUM[287] := '';
   NUM[288] := '';
   NUM[289] := '';
   NUM[290] := '';
   NUM[291] := '';
   NUM[292] := '';
   NUM[293] := '';
   NUM[294] := '';
   NUM[295] := '';
   NUM[296] := '';
   NUM[297] := '';
   NUM[298] := '';
   NUM[299] := '';
   NUM[300] := '';
   NUM[301] := '';
   NUM[302] := '';
   NUM[303] := '';
   NUM[304] := '';
   NUM[305] := '';
   NUM[306] := '';
   NUM[307] := '';
   NUM[308] := '';
   NUM[309] := '';
   NUM[310] := '';
   NUM[311] := '';
   NUM[312] := '';
   NUM[313] := '';
   NUM[314] := '';
   NUM[315] := '';
   NUM[316] := '';
   NUM[317] := '';
   NUM[318] := '';
   NUM[319] := '';
   NUM[320] := '';
   NUM[321] := '';
   NUM[322] := '';
   NUM[323] := '';
   NUM[324] := '';
   NUM[325] := '';
   NUM[326] := '';
   NUM[327] := '';
   NUM[328] := '';
   NUM[329] := '';
   NUM[330] := '';
   NUM[331] := '';
   NUM[332] := '';
   NUM[333] := '';
   NUM[334] := '';
   NUM[335] := '';
   NUM[336] := '';
   NUM[337] := '';
   NUM[338] := '';
   NUM[339] := '';
   NUM[340] := '';
   NUM[341] := '';
   NUM[342] := '';
   NUM[343] := '';
   NUM[344] := '';
   NUM[345] := '';
   NUM[346] := '';
   NUM[347] := '';
   NUM[348] := '';
   NUM[349] := '';
   NUM[350] := '';
   NUM[351] := '';
   NUM[352] := '';
   NUM[353] := '';
   NUM[354] := '';
   NUM[355] := '';
   NUM[356] := '';
   NUM[357] := '';
   NUM[358] := '';
   NUM[359] := '';
   NUM[360] := '';
   NUM[361] := '';
   NUM[362] := '';
   NUM[363] := '';
   NUM[364] := '';
   NUM[365] := '';
   NUM[366] := '';
   NUM[367] := '';
   NUM[368] := '';
   NUM[369] := '';
   NUM[370] := '';
   NUM[371] := '';
   NUM[372] := '';
   NUM[373] := '';
   NUM[374] := '';
   NUM[375] := '';
   NUM[376] := '';
   NUM[377] := '';
   NUM[378] := '';
   NUM[379] := '';
   NUM[380] := '';
   NUM[381] := '';
   NUM[382] := '';
   NUM[383] := '';
   NUM[384] := '';
   NUM[385] := '';
   NUM[386] := '';
   NUM[387] := '';
   NUM[388] := '';
   NUM[389] := '';
   NUM[390] := '';
   NUM[391] := '';
   NUM[392] := '';
   NUM[393] := '';
   NUM[394] := '';
   NUM[395] := '';
   NUM[396] := '';
   NUM[397] := '';
   NUM[398] := '';
   NUM[399] := '';
   NUM[400] := '';
   NUM[401] := '';
   NUM[402] := '';
   NUM[403] := '';
   NUM[404] := '';
   NUM[405] := '';
   NUM[406] := '';
   NUM[407] := '';
   NUM[408] := '';
   NUM[409] := '';
   NUM[410] := '';
   NUM[411] := '';
   NUM[412] := '';
   NUM[413] := '';
   NUM[414] := '';
   NUM[415] := '';
   NUM[416] := '';
   NUM[417] := '';
   NUM[418] := '';
   NUM[419] := '';
   NUM[420] := '';
   NUM[421] := '';
   NUM[422] := '';
   NUM[423] := '';
   NUM[424] := '';
   NUM[425] := '';
   NUM[426] := '';
   NUM[427] := '';
   NUM[428] := '';
   NUM[429] := '';
   NUM[430] := '';
   NUM[431] := '';
   NUM[432] := '';
   NUM[433] := '';
   NUM[434] := '';
   NUM[435] := '';
   NUM[436] := '';
   NUM[437] := '';
   NUM[438] := '';
   NUM[439] := '';
   NUM[440] := '';
   NUM[441] := '';
   NUM[442] := '';
   NUM[443] := '';
   NUM[444] := '';
   NUM[445] := '';
   NUM[446] := '';
   NUM[447] := '';
   NUM[448] := '';
   NUM[449] := '';
   NUM[450] := '';
   NUM[451] := '';
   NUM[452] := '';
   NUM[453] := '';
   NUM[454] := '';
   NUM[455] := '';
   NUM[456] := '';
   NUM[457] := '';
   NUM[458] := '';
   NUM[459] := '';
   NUM[460] := '';
   NUM[461] := '';
   NUM[462] := '';
   NUM[463] := '';
   NUM[464] := '';
   NUM[465] := '';
   NUM[466] := '';
   NUM[467] := '';
   NUM[468] := '';
   NUM[469] := '';
   NUM[470] := '';
   NUM[471] := '';
   NUM[472] := '';
   NUM[473] := '';
   NUM[474] := '';
   NUM[475] := '';
   NUM[476] := '';
   NUM[477] := '';
   NUM[478] := '';
   NUM[479] := '';
   NUM[480] := '';
   NUM[481] := '';
   NUM[482] := '';
   NUM[483] := '';
   NUM[484] := '';
   NUM[485] := '';
   NUM[486] := '';
   NUM[487] := '';
   NUM[488] := '';
   NUM[489] := '';
   NUM[490] := '';
   NUM[491] := '';
   NUM[492] := '';
   NUM[493] := '';
   NUM[494] := '';
   NUM[495] := '';
   NUM[496] := '';
   NUM[497] := '';
   NUM[498] := '';
   NUM[499] := '';
   NUM[500] := '';
   NUM[501] := '';
   NUM[502] := '';
   NUM[503] := '';
   NUM[504] := '';
   NUM[505] := '';
   NUM[506] := '';
   NUM[507] := '';
   NUM[508] := '';
   NUM[509] := '';
   NUM[510] := '';
   NUM[511] := '';
   NUM[512] := '';
   NUM[513] := '';
   NUM[514] := '';
   NUM[515] := '';
   NUM[516] := '';
   NUM[517] := '';
   NUM[518] := '';
   NUM[519] := '';
   NUM[520] := '';
   NUM[521] := '';
   NUM[522] := '';
   NUM[523] := '';
   NUM[524] := '';
   NUM[525] := '';
   NUM[526] := '';
   NUM[527] := '';
   NUM[528] := '';
   NUM[529] := '';
   NUM[530] := '';
   NUM[531] := '';
   NUM[532] := '';
   NUM[533] := '';
   NUM[534] := '';
   NUM[535] := '';
   NUM[536] := '';
   NUM[537] := '';
   NUM[538] := '';
   NUM[539] := '';
   NUM[540] := '';
   NUM[541] := '';
   NUM[542] := '';
   NUM[543] := '';
   NUM[544] := '';
   NUM[545] := '';
   NUM[546] := '';
   NUM[547] := '';
   NUM[548] := '';
   NUM[549] := '';
   NUM[550] := '';
   NUM[551] := '';
   NUM[552] := '';
   NUM[553] := '';
   NUM[554] := '';
   NUM[555] := '';
   NUM[556] := '';
   NUM[557] := '';
   NUM[558] := '';
   NUM[559] := '';
   NUM[560] := '';
   NUM[561] := '';
   NUM[562] := '';
   NUM[563] := '';
   NUM[564] := '';
   NUM[565] := '';
   NUM[566] := '';
   NUM[567] := '';
   NUM[568] := '';
   NUM[569] := '';
   NUM[570] := '';
   NUM[571] := '';
   NUM[572] := '';
   NUM[573] := '';
   NUM[574] := '';
   NUM[575] := '';
   NUM[576] := '';
   NUM[577] := '';
   NUM[578] := '';
   NUM[579] := '';
   NUM[580] := '';
   NUM[581] := '';
   NUM[582] := '';
   NUM[583] := '';
   NUM[584] := '';
   NUM[585] := '';
   NUM[586] := '';
   NUM[587] := '';
   NUM[588] := '';
   NUM[589] := '';
   NUM[590] := '';
   NUM[591] := '';
   NUM[592] := '';
   NUM[593] := '';
   NUM[594] := '';
   NUM[595] := '';
   NUM[596] := '';
   NUM[597] := '';
   NUM[598] := '';
   NUM[599] := '';
   NUM[600] := '';
   NUM[601] := '';
   NUM[602] := '';
   NUM[603] := '';
   NUM[604] := '';
   NUM[605] := '';
   NUM[606] := '';
   NUM[607] := '';

END_DATA_BLOCK
DATA_BLOCK "DI_STRING_NAMES_GER"
{ S7_Optimized_Access := 'FALSE' }
VERSION : 0.1
NON_RETAIN
"DT_DI_STRING_NAMES"

BEGIN
   NUM[0] := 'Wartungsschalter aktiv (-S100)';
   NUM[1] := 'Ortssteuerung aktiv (-S103)';
   NUM[2] := 'Automatische Steuerung aktiv (-S104)';
   NUM[3] := 'Start-Drucktaste gedrueckt (-S210)';
   NUM[4] := 'Stop-Drucktaste gedrueckt (-S211)';
   NUM[5] := 'Alarme zuruecksetzen (-S302)';
   NUM[6] := 'ESD-Drucktaste aktiv (-S301)';
   NUM[7] := 'Externe ESD-Drucktaste aktiv';
   NUM[8] := 'ESD-Relais OK (-K301)';
   NUM[9] := 'Watchdog aktiv';
   NUM[10] := 'Externe Signale PS OK (-F43)';
   NUM[11] := 'DC MCB Gruppenalarm (-F34, -F38, -F40)';
   NUM[12] := 'DC MCB Gruppenausloesung (-F36, -F37, -F39)';
   NUM[13] := 'Synchronisation manuell';
   NUM[14] := 'Synchronisation automatisch';
   NUM[15] := 'Synchronisationsstart';
   NUM[16] := 'Synchronisationsstopp';
   NUM[17] := 'Synchronisationsgeraet OK';
   NUM[18] := 'Synchronisation aktiv (-K1)';
   NUM[19] := 'Synchronisationsgeschwindigkeit runter (-F100)';
   NUM[20] := 'Synchronisationsgeschwindigkeit hoch (-F100)';
   NUM[21] := 'GCB-Schalter EIN-Drucktaste';
   NUM[22] := 'GCB-Schalter AUS-Drucktaste';
   NUM[23] := 'GCB geschlossen (-Q1)';
   NUM[24] := 'GCB offen (-Q1)';
   NUM[25] := 'Generator-Ueberdrehzahlausloesung (-K311)';
   NUM[26] := 'Fernstart';
   NUM[27] := 'Fernstopp';
   NUM[28] := 'Schnellabschaltungsrelais OK (-K401)';
   NUM[29] := 'Reserve 29';
   NUM[30] := 'Synchroskop-Schuetz geschlossen (-K2)';
   NUM[31] := 'Reserve 31';
   NUM[32] := 'AC MCB Gruppenalarm OK';
   NUM[33] := 'AC MCB Gruppenausloesung OK';
   NUM[34] := 'DC MCB Gruppenalarm (-F36)';
   NUM[35] := 'DC MCB Gruppenausloesung (-F38,39,40,44,45)';
   NUM[36] := 'Hauptleistungsschalter EIN (-F1)';
   NUM[37] := 'Hauptleistungsschalter AUS';
   NUM[38] := 'Hauptleistungsschalter manuell';
   NUM[39] := 'Hauptleistungsschalter automatisch';
   NUM[40] := 'Hauptleistungsschalter ausgeloest';
   NUM[41] := 'Diesel-Leistungsschalter EIN';
   NUM[42] := 'Diesel-Leistungsschalter AUS';
   NUM[43] := 'Diesel-Leistungsschalter manuell';
   NUM[44] := 'Diesel-Leistungsschalter automatisch';
   NUM[45] := 'Ueberdrehschutz MCB OK';
   NUM[46] := 'AC-Spannung OK (-F411, -K411)';
   NUM[47] := 'Spannung vor Hauptleistungsschalter OK (-F411, -K411)';
   NUM[48] := 'Spannung vor Diesel-Leistungsschalter OK';
   NUM[49] := 'Ueberspannungsableiter OK (-FU1)';
   NUM[50] := 'AC/DC Gleichrichter 1 OK (-F60, -U101)';
   NUM[51] := 'AC/DC Gleichrichter 2 OK (-F61, -U102)';
   NUM[52] := 'AC/DC Gleichrichter 3 OK';
   NUM[53] := 'Batterie verbunden (-FB, -F421, -K201)';
   NUM[54] := 'Gemeinsame DC-Stromversorgung OK (-F0)';
   NUM[55] := 'Einlass-Schaltschrank AC-Versorgung MCB EIN (-F7)';
   NUM[56] := 'Externe Lasten MCB EIN (-F55,-F56,-F57)';
   NUM[57] := 'Kraftwerksverteilerschrank MCB geschlossen (-F5)';
   NUM[58] := '6,3 MV Schaltanlagensteuerung MCB OK (-F43)';
   NUM[59] := 'Steuerschrank DC-Versorgung MCB geschlossen (-F1';
   NUM[60] := 'GCB-Schaltschrank DC-Versorgung MCB EIN (-F11)';
   NUM[61] := 'MV-Schaltschrank DC-Versorgung MCB geschlossen (';
   NUM[62] := 'AKA01 - MV AC Stromversorgung (-F82)';
   NUM[63] := 'Gemeinsame DC-Stromversorgung (-F0)';
   NUM[64] := 'Reserve 64';
   NUM[65] := 'Reserve 65';
   NUM[66] := 'Reserve 66';
   NUM[67] := 'Reserve 67';
   NUM[68] := 'Netzspannungswandler Messung';
   NUM[69] := 'Gen';
   NUM[70] := 'Reserve 70';
   NUM[71] := 'Reserve 71';
   NUM[72] := 'Reserve 72';
   NUM[73] := 'Reserve 73';
   NUM[74] := 'GCB bereit zum Schliessen (-Q1)';
   NUM[75] := 'Reserve 75';
   NUM[76] := 'GCB-Feder geladen (-Q1)';
   NUM[77] := 'Reserve 77';
   NUM[78] := 'Generator-Leistungsschalter Steuerung MCB EIN (-F62)';
   NUM[79] := 'Reserve 79';
   NUM[80] := 'Reserve 80';
   NUM[81] := 'Reserve 81';
   NUM[82] := 'Reserve 82';
   NUM[83] := 'Ueberspannungsableiter OK (-F60, -FU1)';
   NUM[84] := 'Reserve 84';
   NUM[85] := 'Reserve 85';
   NUM[86] := 'DC Gruppen-Ausloesung (-F4, -F7, -F11, -F14)';
   NUM[87] := 'Hilfstransformator-Versorgungsschalter EIN (-Q2)';
   NUM[88] := 'Reserve 88';
   NUM[89] := 'Ueberspannungsableiter 2 OK (-F61, -FU2)';
   NUM[90] := 'Reserve 90';
   NUM[91] := 'Reserve 91';
   NUM[92] := 'Reserve 92';
   NUM[93] := 'Reserve 93';
   NUM[94] := 'Reserve 94';
   NUM[95] := 'Lampenpruefung (-S203)';
   NUM[96] := 'Generatorspannungsmessung';
   NUM[97] := 'Reserve';
   NUM[98] := 'Reserve';
   NUM[99] := 'Generatorheizung MCB geschlossen (-F53)';
   NUM[100] := 'Generatorheizung Schuetz geschlossen (-K74)';
   NUM[101] := 'Reserve';
   NUM[102] := 'Reserve';
   NUM[103] := 'Reserve';
   NUM[104] := 'Reserve';
   NUM[105] := 'Reserve';
   NUM[106] := 'Reserve';
   NUM[107] := 'Reserve';
   NUM[108] := 'Reserve';
   NUM[109] := 'Reserve';
   NUM[110] := 'Generator Schmieroelstand min';
   NUM[111] := 'Generator Schmierpumpe EIN (-SG24)';
   NUM[112] := 'Generator Vibration Ausloesung (-VSE002)';
   NUM[113] := 'Reserve';
   NUM[114] := 'Reserve';
   NUM[115] := 'Reserve';
   NUM[116] := 'Reserve';
   NUM[117] := 'Reserve';
   NUM[118] := 'Reserve';
   NUM[119] := 'Reserve';
   NUM[120] := 'Reserve';
   NUM[121] := 'Reserve';
   NUM[122] := 'Reserve';
   NUM[123] := 'Reserve';
   NUM[124] := 'Reserve';
   NUM[125] := 'Reserve';
   NUM[126] := 'Reserve';
   NUM[127] := 'Reserve';
   NUM[128] := 'Generator Schutz Ausloesung (-F100)';
   NUM[129] := 'Reserve';
   NUM[130] := 'Reserve';
   NUM[131] := 'Generator Schutz aktiv (-F100)';
   NUM[132] := 'Reserve';
   NUM[133] := 'Reserve';
   NUM[134] := 'Reserve';
   NUM[135] := 'Reserve';
   NUM[136] := 'Reserve';
   NUM[137] := 'Reserve';
   NUM[138] := 'Reserve';
   NUM[139] := 'Reserve';
   NUM[140] := 'AJA04 - Leitungsschutz Ausloesung 1 (-F200)';
   NUM[141] := 'AJA04 - Leitungsschutz Ausloesung 2 (-F200)';
   NUM[142] := 'AJA04 - Leitungsschutz Alarm (-F200)';
   NUM[143] := 'AKA04 - Leitungsschutz aktiv (-F200)';
   NUM[144] := 'Reserve';
   NUM[145] := 'Reserve';
   NUM[146] := 'Reserve';
   NUM[147] := 'Reserve';
   NUM[148] := 'Reserve';
   NUM[149] := 'Reserve';
   NUM[150] := 'Reserve';
   NUM[151] := 'Reserve';
   NUM[152] := 'Reserve';
   NUM[153] := 'Reserve';
   NUM[154] := 'Reserve';
   NUM[155] := 'Reserve';
   NUM[156] := 'Reserve';
   NUM[157] := 'Reserve';
   NUM[158] := 'Reserve';
   NUM[159] := 'Reserve';
   NUM[160] := 'Ueberspannungsableiter OK (-FU1)';
   NUM[161] := 'Stromversorgung CB EIN (-Q1)';
   NUM[162] := 'Gleichrichter OK (-F3)';
   NUM[163] := 'DC MCB OK Gruppenalarm (-F31, -F40)';
   NUM[164] := 'AC MCB OK Gruppenalarm (-F2,-F5,-F6)';
   NUM[165] := 'PSU (-U101) - ALARM';
   NUM[166] := 'PSU (-U101) - Batteriebetrieb';
   NUM[167] := 'PSU (-U101) - Ladebetrieb';
   NUM[168] := 'Reserve';
   NUM[169] := 'Reserve';
   NUM[170] := 'Reserve';
   NUM[171] := 'Reserve';
   NUM[172] := 'Reserve';
   NUM[173] := 'Reserve';
   NUM[174] := 'Reserve';
   NUM[175] := 'Reserve';
   NUM[176] := 'Reserve';
   NUM[177] := 'Reserve';
   NUM[178] := 'Reserve';
   NUM[179] := 'Reserve';
   NUM[180] := 'Reserve';
   NUM[181] := 'Reserve';
   NUM[182] := 'Reserve';
   NUM[183] := 'Reserve';
   NUM[184] := 'Reserve';
   NUM[185] := 'Reserve';
   NUM[186] := 'Reserve';
   NUM[187] := 'Reserve';
   NUM[188] := 'Reserve';
   NUM[189] := 'Reserve';
   NUM[190] := 'Reserve';
   NUM[191] := 'Reserve';
   NUM[192] := 'MIV geschlossen (-1K22)';
   NUM[193] := 'Reserve';
   NUM[194] := 'MIV offen (-1K21)';
   NUM[195] := 'Reserve';
   NUM[196] := 'Reserve';
   NUM[197] := 'MIV CB geschlossen (-F52)';
   NUM[198] := 'MIV Schuetz geschlossen (-K52, -K53)';
   NUM[199] := 'MIV Heizung MCB geschlossen (-F58)';
   NUM[200] := 'Reserve';
   NUM[201] := 'Bypass offen (-ACRON)';
   NUM[202] := 'Bypass geschlossen (-ACRON)';
   NUM[203] := 'Bypass Versorgung MCB EIN (-F40)';
   NUM[204] := 'Reserve';
   NUM[205] := 'Bypass Schuetz geschlossen (-K101,-K102)';
   NUM[206] := 'Bypass oeffnen Schuetz EIN (-K102)';
   NUM[207] := 'Bypass schliessen Schuetz EIN (-K101)';
   NUM[208] := 'Reserve';
   NUM[209] := 'Reserve';
   NUM[210] := 'Reserve';
   NUM[211] := 'Reserve';
   NUM[212] := 'Reserve';
   NUM[213] := 'Reserve';
   NUM[214] := 'MIV Drehmoment-Schalter geschlossen (-1K06)';
   NUM[215] := 'MIV Drehmoment-Schalter offen (-1K05)';
   NUM[216] := 'MIV Thermoschalter (-1K13)';
   NUM[217] := 'Reserve';
   NUM[218] := 'Reserve';
   NUM[219] := 'Reserve';
   NUM[220] := 'Reserve';
   NUM[221] := 'Reserve';
   NUM[222] := 'Reserve';
   NUM[223] := 'Reserve';
   NUM[224] := 'Reserve';
   NUM[225] := 'HPU Leitungsfilter Ausloesung (-600S1)';
   NUM[226] := 'Reserve';
   NUM[227] := 'Reserve';
   NUM[228] := 'Accumulator ESD Druck OK (-640B3)';
   NUM[229] := 'HPU min';
   NUM[230] := 'HPU max';
   NUM[231] := 'Accumulator Start/Stopp Pumpe (-X3)';
   NUM[232] := 'Systemdruck OK (-640B4)';
   NUM[233] := 'HPU Oelstand zu niedrig (-640B2)';
   NUM[234] := 'HPU Oelstand niedrig (-640B2)';
   NUM[235] := 'Reserve';
   NUM[236] := 'HPU Oeltemperatur zu hoch (-640B1)';
   NUM[237] := 'HPU Oeltemperatur hoch (-640B1)';
   NUM[238] := 'Reserve';
   NUM[239] := 'Reserve';
   NUM[240] := 'Reserve';
   NUM[241] := 'Reserve';
   NUM[242] := 'HPU Heizung MCB geschlossen (-F57)';
   NUM[243] := 'HPU Heizung Schuetz geschlossen (-K57)';
   NUM[244] := 'HPU Steuerung MCB geschlossen (-F59)';
   NUM[245] := 'Reserve';
   NUM[246] := 'Reserve';
   NUM[247] := 'Reserve';
   NUM[248] := 'Reserve';
   NUM[249] := 'Reserve';
   NUM[250] := 'Reserve';
   NUM[251] := 'Reserve';
   NUM[252] := 'Reserve';
   NUM[253] := 'Reserve';
   NUM[254] := 'Reserve';
   NUM[255] := 'Reserve';
   NUM[256] := 'Reserve';
   NUM[257] := 'Reserve';
   NUM[258] := 'Reserve';
   NUM[259] := 'HPU Pumpe CB geschlossen (-F51)';
   NUM[260] := 'HPU Pumpe Schuetz geschlossen (-K51)';
   NUM[261] := 'Reserve';
   NUM[262] := 'Reserve';
   NUM[263] := 'Reserve';
   NUM[264] := 'Pumpe 2 MCB EIN (-F2)';
   NUM[265] := 'Pumpe 2 Schuetz EIN (-K2)';
   NUM[266] := 'Reserve';
   NUM[267] := 'Reserve';
   NUM[268] := 'Reserve';
   NUM[269] := 'Reserve';
   NUM[270] := 'Reserve';
   NUM[271] := 'Reserve';
   NUM[272] := 'Reserve';
   NUM[273] := 'Reserve';
   NUM[274] := 'Reserve';
   NUM[275] := 'Reserve';
   NUM[276] := 'Reserve';
   NUM[277] := 'Reserve';
   NUM[278] := 'Reserve';
   NUM[279] := 'Reserve';
   NUM[280] := 'Reserve';
   NUM[281] := 'Reserve';
   NUM[282] := 'Reserve';
   NUM[283] := 'Reserve';
   NUM[284] := 'Reserve';
   NUM[285] := 'Reserve';
   NUM[286] := 'Reserve';
   NUM[287] := 'Reserve';
   NUM[288] := 'Reserve';
   NUM[289] := 'Reserve';
   NUM[290] := 'Reserve';
   NUM[291] := 'Reserve';
   NUM[292] := 'Reserve';
   NUM[293] := 'Reserve';
   NUM[294] := 'Reserve';
   NUM[295] := 'Reserve';
   NUM[296] := 'Reserve';
   NUM[297] := 'Reserve';
   NUM[298] := 'Reserve';
   NUM[299] := 'Reserve';
   NUM[300] := 'Reserve';
   NUM[301] := 'Reserve';
   NUM[302] := 'Reserve';
   NUM[303] := 'Reserve';
   NUM[304] := 'Reserve';
   NUM[305] := 'Reserve';
   NUM[306] := 'Reserve';
   NUM[307] := 'Reserve';
   NUM[308] := 'Reserve';
   NUM[309] := 'Reserve';
   NUM[310] := 'Reserve';
   NUM[311] := 'Reserve';
   NUM[312] := 'Reserve';
   NUM[313] := 'Reserve';
   NUM[314] := 'Reserve';
   NUM[315] := 'Reserve';
   NUM[316] := 'Reserve';
   NUM[317] := 'Reserve';
   NUM[318] := 'Reserve';
   NUM[319] := 'Reserve';
   NUM[320] := 'Reserve';
   NUM[321] := 'Reserve';
   NUM[322] := 'Reserve';
   NUM[323] := 'Reserve';
   NUM[324] := 'Reserve';
   NUM[325] := 'Reserve';
   NUM[326] := 'Reserve';
   NUM[327] := 'Reserve';
   NUM[328] := 'Reserve';
   NUM[329] := 'Reserve';
   NUM[330] := 'Reserve';
   NUM[331] := 'Reserve';
   NUM[332] := 'Reserve';
   NUM[333] := 'Reserve';
   NUM[334] := 'Reserve';
   NUM[335] := 'Reserve';
   NUM[336] := 'Reserve';
   NUM[337] := 'Reserve';
   NUM[338] := 'Reserve';
   NUM[339] := 'Reserve';
   NUM[340] := 'Reserve';
   NUM[341] := 'Reserve';
   NUM[342] := 'Reserve';
   NUM[343] := 'Reserve';
   NUM[344] := 'Reserve';
   NUM[345] := 'Reserve';
   NUM[346] := 'Reserve';
   NUM[347] := 'Reserve';
   NUM[348] := 'Reserve';
   NUM[349] := 'Reserve';
   NUM[350] := 'Reserve';
   NUM[351] := 'Reserve';
   NUM[352] := 'Reserve';
   NUM[353] := 'Reserve';
   NUM[354] := 'Heizung der Laufschaufeln MCB EIN (-F54)';
   NUM[355] := 'Antrieb der Laufschaufeln Steuerung';
   NUM[356] := 'Antrieb der Laufschaufeln Steuerung';
   NUM[357] := 'Heizung des Schutzes MCB EIN (-F49)';
   NUM[358] := 'Antrieb der Laufschaufeln CB EIN (-F51)';
   NUM[359] := 'Antrieb des Schutzes CB EIN (-F47)';
   NUM[360] := 'Antrieb des Schutzes Steuerung';
   NUM[361] := 'Antrieb des Schutzes Steuerung';
   NUM[362] := 'Heizung des Schutzes Steuerung';
   NUM[363] := 'Uberdrehzahl-Abschaltung (Turbine) (-K312)';
   NUM[364] := 'Drehmoment-Schalter des Schutzes "C"';
   NUM[365] := 'Drehmoment-Schalter des Schutzes "O"';
   NUM[366] := 'Endschalter des Schutzes "C"';
   NUM[367] := 'Endschalter des Schutzes "O"';
   NUM[368] := 'Drehmoment-Schalter der Laufschaufeln "C"';
   NUM[369] := 'Drehmoment-Schalter der Laufschaufeln "O"';
   NUM[370] := 'Endschalter der Laufschaufeln "C"';
   NUM[371] := 'Endschalter der Laufschaufeln "O"';
   NUM[372] := 'Thermoschalter der Laufschaufeln (-1K11)';
   NUM[373] := 'Reserve';
   NUM[374] := 'Reserve';
   NUM[375] := 'Reserve';
   NUM[376] := 'Reserve';
   NUM[377] := 'Reserve';
   NUM[378] := 'Reserve';
   NUM[379] := 'Reserve';
   NUM[380] := 'Reserve';
   NUM[381] := 'Reserve';
   NUM[382] := 'Reserve';
   NUM[383] := 'Reserve';
   NUM[384] := 'Einheitstrafo 1BAT10 - Temperaturalarm (-1K37)';
   NUM[385] := 'Einheitstrafo 1BAT10 - Temperatur-Abschaltung (-';
   NUM[386] := 'Transformator - Druckalarm (-1K01)';
   NUM[387] := 'Einheitstrafo 1BAT10 - Druck-Abschaltung (-1K36)';
   NUM[388] := 'Reserve';
   NUM[389] := 'Reserve';
   NUM[390] := 'Einheitstrafo - Buchholz-Alarm';
   NUM[391] := 'Einheitstrafo 1BAT10 - Gas-Abschaltung (-1K35)';
   NUM[392] := 'Reserve';
   NUM[393] := 'Reserve';
   NUM[394] := 'Reserve';
   NUM[395] := 'Reserve';
   NUM[396] := 'Reserve';
   NUM[397] := 'Reserve';
   NUM[398] := 'Reserve';
   NUM[399] := 'Reserve';
   NUM[400] := 'Reserve';
   NUM[401] := 'Reserve';
   NUM[402] := 'Reserve';
   NUM[403] := 'Reserve';
   NUM[404] := 'Reserve';
   NUM[405] := 'Reserve';
   NUM[406] := 'Reserve';
   NUM[407] := 'Reserve';
   NUM[408] := 'Reserve';
   NUM[409] := 'Reserve';
   NUM[410] := 'Reserve';
   NUM[411] := 'Reserve';
   NUM[412] := 'Reserve';
   NUM[413] := 'SS trafo - Wickeltemperatur U Ok (-TH145)';
   NUM[414] := 'SS trafo - Wickeltemperatur V Ok (-TH145)';
   NUM[415] := 'SS trafo - Wickeltemperatur W Ok (-TH145)';
   NUM[416] := 'Reserve';
   NUM[417] := 'Reserve';
   NUM[418] := 'Reserve';
   NUM[419] := 'Reserve';
   NUM[420] := 'Reserve';
   NUM[421] := 'Reserve';
   NUM[422] := 'Reserve';
   NUM[423] := 'Reserve';
   NUM[424] := 'Reserve';
   NUM[425] := 'Reserve';
   NUM[426] := 'Reserve';
   NUM[427] := 'Reserve';
   NUM[428] := 'Reserve';
   NUM[429] := 'Reserve';
   NUM[430] := 'Reserve';
   NUM[431] := 'Reserve';
   NUM[432] := 'Reserve';
   NUM[433] := 'Reserve';
   NUM[434] := 'Reserve';
   NUM[435] := 'Reserve';
   NUM[436] := 'Reserve';
   NUM[437] := 'Reserve';
   NUM[438] := 'Reserve';
   NUM[439] := 'Reserve';
   NUM[440] := 'Reserve';
   NUM[441] := 'Reserve';
   NUM[442] := 'Reserve';
   NUM[443] := 'Reserve';
   NUM[444] := 'Reserve';
   NUM[445] := 'Reserve';
   NUM[446] := 'Reserve';
   NUM[447] := 'Reserve';
   NUM[448] := 'Anlaufkontakt geschlossen (-K1)';
   NUM[449] := 'Synchronisation Spannung niedriger (-F100)';
   NUM[450] := 'Synchronisation Spannung hoher (-F100)';
   NUM[451] := 'Anregungsgerat Abschaltung (DV0 - RLY1)';
   NUM[452] := 'Anregungsalarm (DECS - AL2, -1K13)';
   NUM[453] := 'Anregungsdiode Uberwachung Abschaltung (DV0 - RL';
   NUM[454] := 'AVR Relais 1';
   NUM[455] := 'AVR Relais 2';
   NUM[456] := 'Reserve';
   NUM[457] := 'AVR Watchdog OK (-K111)';
   NUM[458] := 'AVR nicht abgeschaltet (-K112)';
   NUM[459] := 'AVR Start';
   NUM[460] := 'AVR Begrenzung Aktiv';
   NUM[461] := 'Reserve';
   NUM[462] := 'Reserve';
   NUM[463] := 'Reserve';
   NUM[464] := 'AVR DO 1';
   NUM[465] := 'AVR DO 2';
   NUM[466] := 'AVR DO 3';
   NUM[467] := 'EXC AREP PS OK (-Q1)';
   NUM[468] := 'Reserve';
   NUM[469] := 'Reserve';
   NUM[470] := 'Reserve';
   NUM[471] := 'Reserve';
   NUM[472] := 'Reserve';
   NUM[473] := 'Reserve';
   NUM[474] := 'Reserve';
   NUM[475] := 'Reserve';
   NUM[476] := 'Reserve';
   NUM[477] := 'Reserve';
   NUM[478] := 'Reserve';
   NUM[479] := 'Reserve';
   NUM[480] := '0AKA01 - Trennschalter geschlossen (-Q2)';
   NUM[481] := '0AKA01 - Trennschalter geoffnet (-Q2)';
   NUM[482] := 'Reserve';
   NUM[483] := '0AKA01 - Erdungsschalter geschlossen (-Q3)';
   NUM[484] := '0AKA01 - Erdungsschalter geoffnet (-Q3)';
   NUM[485] := '0AKA01 - Spannungsuberwachungsrelais geschlossen';
   NUM[486] := '0AKA02 - Spannungs-Trafo MCB geschlossen (-Q11)';
   NUM[487] := '0AKA01 - CB Feder geladen (-Q0)';
   NUM[488] := 'Reserve';
   NUM[489] := '0AKA01 - Fernsteuerung (-S60)';
   NUM[490] := '0AKA01 - Leistungsschalter geschlossen (-Q1)';
   NUM[491] := '0AKA01 - Leistungsschalter geoffnet (-Q1)';
   NUM[492] := 'Reserve';
   NUM[493] := 'Reserve';
   NUM[494] := '0AKA01 - DC MCB OK Gruppe 1 Abschaltung (-F14)';
   NUM[495] := '0AKA01 - Gasdruck OK (-Q1)';
   NUM[496] := 'Hebel eingesetzt';
   NUM[497] := '0AKA01 - 2. Shuntfreigabe MCB EIN (-F5)';
   NUM[498] := 'Reserve';
   NUM[499] := '0AKA01 - DC Steuerung und Signal';
   NUM[500] := '0AKA01 - AC Steuerung und Signal';
   NUM[501] := '0AKA01 - Ladegerat MCB geschlossen (-Q5)';
   NUM[502] := '0AGA02 - Ausgangsleitung CB Dienst';
   NUM[503] := '0AKA01 - MV Heizungen EIN (-Q6)';
   NUM[504] := 'Reserve';
   NUM[505] := 'Reserve';
   NUM[506] := 'Reserve';
   NUM[507] := 'Reserve';
   NUM[508] := 'Reserve';
   NUM[509] := 'Reserve';
   NUM[510] := 'Reserve';
   NUM[511] := 'Reserve';
   NUM[512] := 'AJA04 - DS geschlossen (-Q2)';
   NUM[513] := 'AJA04 - DS geoffnet (-Q2)';
   NUM[514] := 'Reserve';
   NUM[515] := 'AJA04 - ES geschlossen (-Q2)';
   NUM[516] := 'AJA04 - ES geoffnet (-Q2)';
   NUM[517] := '0AKA03 - Spannung vorhanden (-F23 -> R1,R2)';
   NUM[518] := 'Reserve';
   NUM[519] := 'Reserve';
   NUM[520] := 'Reserve';
   NUM[521] := 'AJA04 - Lokale Steuerung (-S60)';
   NUM[522] := 'AJA04 - CB geschlossen (-Q1)';
   NUM[523] := 'AJA04 - CB geoffnet (-Q1)';
   NUM[524] := 'Reserve';
   NUM[525] := 'Reserve';
   NUM[526] := 'Reserve';
   NUM[527] := 'Reserve';
   NUM[528] := 'Reserve';
   NUM[529] := 'Reserve';
   NUM[530] := 'Reserve';
   NUM[531] := 'Reserve';
   NUM[532] := 'Reserve';
   NUM[533] := 'Reserve';
   NUM[534] := 'Reserve';
   NUM[535] := 'Reserve';
   NUM[536] := 'Reserve';
   NUM[537] := 'Steuerung und Signal';
   NUM[538] := 'Ladegerat MCB geschlossen (-Q5)';
   NUM[539] := 'Reserve';
   NUM[540] := '0AKA03 - Spannungs-Trafo MCB geschlossen (-Q11)';
   NUM[541] := 'Reserve';
   NUM[542] := 'Reserve';
   NUM[543] := 'Reserve';
   NUM[544] := 'S';
   NUM[545] := 'S';
   NUM[546] := 'S';
   NUM[547] := 'S';
   NUM[548] := 'S';
   NUM[549] := 'S';
   NUM[550] := 'Reserve';
   NUM[551] := 'Reserve';
   NUM[552] := 'Reserve';
   NUM[553] := 'Reserve';
   NUM[554] := 'Reserve';
   NUM[555] := 'Reserve';
   NUM[556] := 'Reserve';
   NUM[557] := 'Reserve';
   NUM[558] := 'Reserve';
   NUM[559] := 'Reserve';
   NUM[560] := 'Reserve';
   NUM[561] := 'Reserve';
   NUM[562] := 'Reserve';
   NUM[563] := 'Reserve';
   NUM[564] := 'Reserve';
   NUM[565] := 'Reserve';
   NUM[566] := 'Reserve';
   NUM[567] := 'Reserve';
   NUM[568] := 'Reserve';
   NUM[569] := 'Reserve';
   NUM[570] := 'Reserve';
   NUM[571] := 'Reserve';
   NUM[572] := 'Reserve';
   NUM[573] := 'Reserve';
   NUM[574] := 'Reserve';
   NUM[575] := 'Reserve';
   NUM[576] := '0AKA03 - CB geoeffnet (-Q1)';
   NUM[577] := '0AKA03 - CB geschlossen (-Q1)';
   NUM[578] := 'Transformator - ausgehende Feder geladen';
   NUM[579] := '0AKA03 - ES geschlossen (-Q3)';
   NUM[580] := '0AKA03 - DS geoeffnet (-Q2)';
   NUM[581] := '0AKA03 - DS geschlossen (-Q2)';
   NUM[582] := 'Transformator - ausgehende Steuerung MCB geschlossen';
   NUM[583] := 'Transformator - ausgehend';
   NUM[584] := '0AKA03 - CB Schliessung (-S60)';
   NUM[585] := '0AKA03 - Steuerung und Signal';
   NUM[586] := '0AKA03 - Ladegeraet MCB geschlossen (-Q5)';
   NUM[587] := 'Transformator - eingehender AC MCB geschlossen';
   NUM[588] := '0AKA03 - Spannungs-Trafo MCB geschlossen (-Q11)';
   NUM[589] := '0AGA01 - VT2 MCB geschlossen';
   NUM[590] := '0AGA01 - VT3 MCB geschlossen';
   NUM[591] := '0AKA03 - ES geoeffnet (-Q3)';
   NUM[592] := '0AKA03 - Spannungsueberwachungsrelais geschlossen (-F23)';
   NUM[593] := 'RESERVE';
   NUM[594] := 'RESERVE';
   NUM[595] := 'RESERVE';
   NUM[596] := 'RESERVE';
   NUM[597] := 'RESERVE';
   NUM[598] := 'RESERVE';
   NUM[599] := 'RESERVE';
   NUM[600] := 'RESERVE';
   NUM[601] := 'RESERVE';
   NUM[602] := 'RESERVE';
   NUM[603] := 'RESERVE';
   NUM[604] := 'RESERVE';
   NUM[605] := 'RESERVE';
   NUM[606] := 'RESERVE';
   NUM[607] := 'RESERVE';

END_DATA_BLOCK
